Fanuc KAREL source: kt00450.KL

-- PROVISIONAL review KL for V1013-1; original PC SHA256 a20fa81160ab018418ff0bc058a59542a3789334beda86828b3b9a5860ec88de
-- Incomplete behavior may be omitted. Consult companion uncertainty JSON. Do not deploy.
PROGRAM KT00450
%NOLOCKGROUP
VAR
  OUT : BOOLEAN
-- UNRESOLVED_DECL Y1 type=002018
-- UNRESOLVED_DECL H2 type=002017
BEGIN
  -- UNRESOLVED_PC offsets 5-19; opcodes 2E,22,9D,33,B2
  -- UNRESOLVED_PC offsets 24-38; opcodes 2E,22,9D,33,B4
  -- UNRESOLVED_PC offsets 43-68; opcodes 22,9D,33,B1,22,9D,33,B3,5C,23
  -- UNRESOLVED_PC offsets 73-77; opcodes 7F
END KT00450
